(* IEC 61131-3 sources: JingjiangMoonbox/Application/Application/任务列表/TensionTask/电机运动/MotionCtl_GantryTrap/HandWheelCtl, 6 files *)

(* ---- StHandWheel.st ---- *)
(*@CES
Name=StHandWheel
Type=Gvl
TypeGuid=2db5746d-d284-4425-9f7f-2663a34b0ebc
Guid=e24024ef-b057-4603-89fd-c6f3dc30d212
HasDeclaration=True
HasImplementation=False
*)
{DECLARATION}
{attribute 'pack_mode' := '1'}
TYPE StHandWheel :
STRUCT
	wButton_HardWheel: WORD;(*手轮按键bit0-bit12对应按键1-13（手轮从左到右，从上到下）*)
// 	byRate_HardWheel: BYTE;(*倍率选择=13：X1;=14：X10;=15：X100;=16：X1000;=26：未定义（1000X后面还有一个档位）*)
// 	byAxisId_HardWheelCtl: BYTE;(*手轮旋钮当前选择
// 								=6：OFF
// 								=17：X
// 								=18：Y
// 								=19：Z
// 								=20：A*)

//2023.9.25.131020|手轮实际是倍率和轴选不是之前的定义，我们交换了一些2023.9.25.13110|
	byKnob_Right: BYTE;(*右选择=13：0档位;
								=14：1档位;
								=15：2档位;
								=16：3档位;
								=26：4档位（1000X后面还有一个档位）*)
	byKnob_Left: BYTE;(*左旋钮当前选择
								=6：0档位
								=17：1档位
								=18：2档位
								=19：3档位
								=20：4档位*)
	lrTargetPos_HardWheel: LREAL;(*当前手轮值-可以通过GT_RN_ZeroHandPos指令清除*)
	byHandWheelSts: BYTE;(**)
	asDisplay_HardWheel_HMI: ARRAY [1..4] OF STRING(16);(*手轮HMI显示-*)
	(*屏显功能说明：
	1.显示信号、电池电量
	2.当前操作色组号、当前操作的轴、标定模式以及标定轴、步进值
	3.显示版辊两侧电机实时位置(mm)
	4.显示网辊两侧电机实时位置(mm)
	(屏显格式说明：1行显示11个字符
	2/3/4行能显示16个字符)*)
	//2024.3.13.142250用于通讯给从站的变量
	arPos_HandWheel: ARRAY [1..4] OF REAL;//4个压力电机位置版辊M-G，网辊M-G
	byCtlId_HandWheel: BYTE;
	byCtlSts_HandWheel: BYTE;
						(*
							bit0:锁定模式
							bit1:运行模式
							bit2:标定DEBUG
							bit3:急停
							bit4:报警
							bit5:版/网切换
							bit6:清零处理
			2025.04.02.144750
							bit7:切换色组
						*)
END_STRUCT
END_TYPE

{IMPLEMENTATION}

(* ---- StHandWheel_BtnCtl.st ---- *)
(*@CES
Name=StHandWheel_BtnCtl
Type=Gvl
TypeGuid=2db5746d-d284-4425-9f7f-2663a34b0ebc
Guid=b84cb397-2bed-4490-8555-fa94b8c7b26f
HasDeclaration=True
HasImplementation=False
*)
{DECLARATION}
TYPE StHandWheel_BtnCtl :
STRUCT
	xReq_Inch_Net: BOOL;//匀墨
	xReqSwitch_Calib: BOOL;
	xReq_Confirm_Adjust_PressDn: BOOL;//位置矫正
	lrPos_HandWheelChange: LREAL;//手轮变化量

	xReqMove_M: BOOL;
	xReqMove_G: BOOL;
	xReqMoveUp: BOOL;
	xReqMoveDn: BOOL;

	xAdjust_V_Up : BOOL;
	xAdjust_V_Dn : BOOL;
	xAdjust_H_M : BOOL;
	xAdjust_H_G : BOOL;

//下面是需要区分版辊压力、网棍压力、张带辊压力的
	axReqLoad_Unload: ARRAY [1..gc_iMax_PressureRoller_Unit] OF BOOL;
	axReqPress_Up: ARRAY [1..gc_iMax_PressureRoller_Unit] OF BOOL;
	axReqPress_Dn: ARRAY [1..gc_iMax_PressureRoller_Unit] OF BOOL;

	axReqMoveFor: ARRAY [1..gc_iMax_PressureRoller_Unit] OF BOOL;
	axReqMoveRev: ARRAY [1..gc_iMax_PressureRoller_Unit] OF BOOL;

	axReq_Confirm_Load_Unload: ARRAY [1..gc_iMax_PressureRoller_Unit] OF BOOL;
	axReq_Confirm_press_up: ARRAY [1..gc_iMax_PressureRoller_Unit] OF BOOL;
	axReq_Confirm_press_dn: ARRAY [1..gc_iMax_PressureRoller_Unit] OF BOOL;

	axFlag_Ctl_Roller_All: ARRAY [1..gc_iMax_PressureRoller_Unit] OF BOOL;//控制的是同进同退-版辊
	axFlag_Ctl_Roller_M: ARRAY [1..gc_iMax_PressureRoller_Unit] OF BOOL;
	axFlag_Ctl_Roller_G: ARRAY [1..gc_iMax_PressureRoller_Unit] OF BOOL;

END_STRUCT
END_TYPE

{IMPLEMENTATION}

(* ---- KS_FB_HandwheelCtl.st ---- *)
(*@CES
Name=KS_FB_HandwheelCtl
Type=FunctionBlock
TypeGuid=6f9dac99-8de1-4efc-8465-68ac443b7d08
Guid=2f871db0-86b8-4868-b4d6-3d54ec95653d
HasDeclaration=True
HasImplementation=True
*)
{DECLARATION}
FUNCTION_BLOCK KS_FB_HandwheelCtl
VAR_INPUT
	i_xEn: BOOL;
	i_byUnitNumMax: BYTE;//色组数
	i_pastStHandWheel: POINTER TO ARRAY [1..MAX_UNIT_NUM] OF StHandWheel;
	i_pastStHandWheel_BtnCtl: POINTER TO ARRAY [1..MAX_UNIT_NUM] OF StHandWheel_BtnCtl;

	i_pabyUnitId_Ctl: POINTER TO ARRAY [1..MAX_UNIT_NUM] OF BYTE;//每个手持器控制的色组，可调整
	i_xFlag_Stop: BOOL;//停机状态
	i_xDebugMode: BOOL;//调试模式
	i_paxNeedZeroPos:  POINTER TO ARRAY [1..MAX_UNIT_NUM] OF BOOL;//手轮计数清零标志
	i_paxFlag_Mode_Calid: POINTER TO ARRAY [1..MAX_UNIT_NUM] OF BOOL;//手持器标定标值
	i_paxFlag_LockHandwheel: POINTER TO ARRAY [1..MAX_UNIT_NUM] OF BOOL;//手持器suoding
	//i_paxFlag_Ctl_Prn: POINTER TO ARRAY [1..MAX_UNIT_NUM] OF BOOL;
	i_paxEn_HandWheel: POINTER TO  ARRAY [1..MAX_UNIT_NUM] OF BOOL;
	i_paxAdjust_Auto_V: POINTER TO  ARRAY [1..MAX_UNIT_NUM] OF BOOL;
	i_paxAdjust_Auto_H: POINTER TO  ARRAY [1..MAX_UNIT_NUM] OF BOOL;

	i_paxAcc_UnitId : POINTER TO  ARRAY [1..MAX_UNIT_NUM] OF BOOL;
END_VAR
VAR_OUTPUT
END_VAR
VAR
	iN: INT;
	iM: INT;
	iRtn : INT;
	xFlag_Handwheel_Unit_One: BOOL;//手持器与色组一对一标值
	axFlag_LockHandwheel: ARRAY [1..MAX_UNIT_NUM] OF BOOL;//手持器锁定标值
	xInit: BOOL:= FALSE;//初始化一些东西
	astStHandWheel_Rec: ARRAY [1..MAX_UNIT_NUM] OF StHandWheel;
	aiCtlStep_Handwheel: ARRAY [1..MAX_UNIT_NUM] OF INT;//手持器锁定标值
	aiCtlUnit_Handwheel: ARRAY [1..MAX_UNIT_NUM] OF INT;//手持器锁定标值
	iTemp:INT:=1;
	aiStartUnitId:ARRAY [1..MAX_UNIT_NUM] OF INT;//非一对一手持器，每个手持器控制的起始
	aiStopUnitId:ARRAY [1..MAX_UNIT_NUM] OF INT;//非一对一手持器，每个手持器控制的结束色组号
	axFlag_Mode_Calid: ARRAY [1..MAX_UNIT_NUM] OF BOOL;//手持器标定标值
	iTimeCnt_Lock:INT:= 600;//超过600个周期没操作，认为可以锁定手轮了防止误操作
	iTimeCnt_Lock_Init:INT:= 3429;//超过600个周期没操作(2分钟)，手轮初始化一次防止进入休眠
	aiCnt_Lock_Num: ARRAY [1..MAX_UNIT_NUM] OF INT;
	aiCnt_Lock_Num_Init: ARRAY [1..MAX_UNIT_NUM] OF INT;
	axFlag_Lock: ARRAY [1..MAX_UNIT_NUM,1..5] OF BOOL;//手轮无动作标志
	iUnitIdCtl: INT;
	aiCnt_LockBtn: ARRAY [1..MAX_UNIT_NUM] OF INT;
	iTimeCnt_LockBtn:INT:= 20;//超过20个周期没操作，认为可以锁定手轮了防止误操作
	afbAcc_AxisId: ARRAY [1..MAX_UNIT_NUM] OF R_TRIG;
	afbDec_AxisId: ARRAY [1..MAX_UNIT_NUM] OF R_TRIG;
	abyAxisId_handwheel: ARRAY [1..MAX_UNIT_NUM] OF BYTE;
	axEn_HandWheel: ARRAY [1..MAX_UNIT_NUM] OF BOOL;
	iK: INT;
	afbTRIG_Switch_Calib: ARRAY [1..MAX_UNIT_NUM] OF R_TRIG;
	fbKS_FB_HandwheelCtl_Reset : KS_FB_HandwheelCtl_Reset;
	xFlag_En_ModeCalib : BOOL;
//2024.12.05.170136 | bai.zy
	xHandWheelCtlSignalUnit : BOOL;
	iHandWheelCount : INT;

	aiAccCtlUnitId_Handwheel: ARRAY [1..MAX_UNIT_NUM] OF INT;//切换色组时手持器锁定的色组号
END_VAR

{IMPLEMENTATION}
IF i_xEn THEN
	IF (i_byUnitNumMax>=1 AND i_byUnitNumMax<= MAX_UNIT_NUM) AND
		i_pastStHandWheel<>0 AND
		i_pabyUnitId_Ctl<>0 AND
		i_pastStHandWheel_BtnCtl <> 0 AND
		i_paxNeedZeroPos <> 0 AND
		i_paxFlag_Mode_Calid <> 0 AND
		i_paxEn_HandWheel <> 0 AND
		i_paxAdjust_Auto_V <> 0 AND
		i_paxAdjust_Auto_H <> 0 THEN

	//	i_pastStHandWheel^[2] := i_pastStHandWheel^[3];
		IF NOT xInit THEN
			xInit:= TRUE;
			FOR iN:=1 TO MAX_UNIT_NUM BY 1 DO
				axFlag_LockHandwheel[iN]:= TRUE;
				axFlag_Mode_Calid[iN]:= FALSE;
				FOR iM:=1 TO 5 BY 1 DO
					axFlag_Lock[iN,iM]:= FALSE;//用于判断手持器无动作的标志
				END_FOR
				aiCtlUnit_Handwheel[iN]:= MAX_UNIT_NUM;
				axEn_HandWheel[iN]:= FALSE;
			END_FOR

		ELSE//初始化完成就可以处理其他了
//2024.3.13.141555
// axEn_HandWheel[1]:= TRUE;
// axEn_HandWheel[2]:= FALSE;
			iHandWheelCount := 0;
			FOR iN := 1 TO i_byUnitNumMax BY 1 DO
				axEn_HandWheel[iN] := i_paxEn_HandWheel^[iN];
				IF axEn_HandWheel[iN] THEN
					iHandWheelCount := iHandWheelCount + 1;
				END_IF
			END_FOR

			IF iHandWheelCount = i_byUnitNumMax THEN
				xHandWheelCtlSignalUnit := TRUE;
			ELSE
				xHandWheelCtlSignalUnit := FALSE;
			END_IF

			FOR iN:=1 TO MAX_UNIT_NUM BY 1 DO
				IF axFlag_LockHandwheel[iN]  OR (NOT axEn_HandWheel[iN]) THEN
					aiCtlStep_Handwheel[iN]:= 1;//锁定状态
				ELSE
					IF xFlag_En_ModeCalib THEN//标定模式2023.7.26.094141更新轴选旋钮，先这么试一下
						IF i_xFlag_Stop AND i_xDebugMode THEN
							axFlag_Mode_Calid[aiCtlUnit_Handwheel[iN]]:= TRUE;
						ELSE
							axFlag_Mode_Calid[aiCtlUnit_Handwheel[iN]]:= FALSE;
							xFlag_En_ModeCalib := FALSE;
						END_IF
 					ELSE
 						axFlag_Mode_Calid[aiCtlUnit_Handwheel[iN]]:= FALSE;
 					END_IF

					IF axFlag_Mode_Calid[aiCtlUnit_Handwheel[iN]] THEN
						aiCtlStep_Handwheel[iN]:= 2;//标定模式
					ELSE
						aiCtlStep_Handwheel[iN]:= 3;//运行模式
					END_IF
				END_IF

			END_FOR
			//换一下吧2024.3.13.132259循环手轮数不好处理

			FOR iN:=1 TO i_byUnitNumMax BY 1 DO
//			FOR iN:=1 TO i_byHandWheel_Num BY 1 DO
				IF i_pastStHandWheel^[iN].wButton_HardWheel=0 THEN//无按钮按下
					axFlag_Lock[iN,1]:= TRUE;
				ELSE
					axFlag_Lock[iN,1]:= FALSE;
				END_IF
				IF i_pastStHandWheel^[iN].byKnob_Left-astStHandWheel_Rec[iN].byKnob_Left=0 THEN//轴选未操作
					axFlag_Lock[iN,2]:= TRUE;
				ELSE
					axFlag_Lock[iN,2]:= FALSE;
				END_IF
				IF i_pastStHandWheel^[iN].byKnob_Right-astStHandWheel_Rec[iN].byKnob_Right=0 THEN//右旋钮无动作
					axFlag_Lock[iN,3]:= TRUE;
				ELSE
					axFlag_Lock[iN,3]:= FALSE;
				END_IF
				IF i_pastStHandWheel^[iN].lrTargetPos_HardWheel-astStHandWheel_Rec[iN].lrTargetPos_HardWheel=0 THEN//手轮无动作
					axFlag_Lock[iN,4]:= TRUE;
				ELSE
					axFlag_Lock[iN,4]:= FALSE;
				END_IF
				IF axFlag_Lock[iN,1] AND axFlag_Lock[iN,2] AND axFlag_Lock[iN,3] AND axFlag_Lock[iN,4] THEN//手轮本周期无动作
					aiCnt_Lock_Num[iN]:= aiCnt_Lock_Num[iN]+1;
					aiCnt_Lock_Num_Init[iN] := aiCnt_Lock_Num_Init[iN] +1;
					IF aiCnt_Lock_Num[iN]>=iTimeCnt_Lock THEN//手持器持续600周期无动作-20s-进入锁定状态
						axFlag_LockHandwheel[iN]:= TRUE;
						aiCnt_Lock_Num[iN] := 0;
					END_IF
					IF aiCnt_Lock_Num_Init[iN]>= iTimeCnt_Lock_Init THEN
;//						iRtn := GT_RN_UsbInit();
						aiCnt_Lock_Num_Init[iN] := 0;
					END_IF
				ELSE
					aiCnt_Lock_Num[iN]:= 0;
					aiCnt_Lock_Num_Init[iN] := 0;
				END_IF

			END_FOR

			FOR iN:=1 TO i_byUnitNumMax BY 1 DO
//			FOR iN:=1 TO i_byHandWheel_Num BY 1 DO
				IF axEn_HandWheel[iN] THEN
					iUnitIdCtl:= aiCtlUnit_Handwheel[iN];
					afbAcc_AxisId[iN](CLK:= i_pastStHandWheel^[iN].wButton_HardWheel.0);
					afbDec_AxisId[iN](CLK:= i_pastStHandWheel^[iN].wButton_HardWheel.1);
					IF abyAxisId_handwheel[iN]<>i_pastStHandWheel^[iN].byKnob_Right THEN
						i_paxNeedZeroPos^[iN]:= TRUE;
						astStHandWheel_Rec[iN].lrTargetPos_HardWheel:= 0;//手轮值清零-好处理
						i_pastStHandWheel^[iN].lrTargetPos_HardWheel:= 0;
					END_IF
					abyAxisId_handwheel[iN]:= i_pastStHandWheel^[iN].byKnob_Right;
					CASE aiCtlStep_Handwheel[iN] OF
						1: //手轮锁定，不允许操作
						//锁定后，所有按钮输入不响应
							IF NOT i_paxAcc_UnitId^[iN] THEN
								IF i_pastStHandWheel^[iN].wButton_HardWheel.0 AND i_pastStHandWheel^[iN].wButton_HardWheel.11 THEN
									//两个按钮同时按下，就认为需要解锁
									axFlag_LockHandwheel[iN]:= FALSE;//解锁
									i_paxNeedZeroPos^[iN]:= TRUE;
									astStHandWheel_Rec[iN].lrTargetPos_HardWheel:= 0;//手轮值清零-好处理
									i_pastStHandWheel^[iN].lrTargetPos_HardWheel:= 0;

								END_IF
							ELSE
								IF afbAcc_AxisId[iN].Q THEN//继续增加
									iUnitIdCtl:= iUnitIdCtl+1;
									FOR iK:=1 TO i_byUnitNumMax BY 1 DO
										IF axEn_HandWheel[iK] THEN
											IF iUnitIdCtl= aiCtlUnit_Handwheel[iK] OR iUnitIdCtl > i_byUnitNumMax THEN//不能与其他手轮冲突
												IF iUnitIdCtl+1 > i_byUnitNumMax THEN//2024.12.05.133431 | bai.zy | 双手轮冲突、超过两个要重新做
													iUnitIdCtl:= 1;
												ELSE
													iUnitIdCtl:= iUnitIdCtl+1;
												END_IF
											END_IF
										END_IF
									END_FOR
									IF iUnitIdCtl>i_byUnitNumMax THEN
										iUnitIdCtl:= 1;
									END_IF
	// 								i_paxAcc_UnitId^[iN] := FALSE;
	// 								axFlag_LockHandwheel[iN]:= FALSE;//解锁
									i_paxNeedZeroPos^[iN]:= TRUE;
									astStHandWheel_Rec[iN].lrTargetPos_HardWheel:= 0;//手轮值清零-好处理
									i_pastStHandWheel^[iN].lrTargetPos_HardWheel:= 0;

									aiCtlUnit_Handwheel[iN]:=iUnitIdCtl;
								ELSIF i_pastStHandWheel^[iN].wButton_HardWheel.1 THEN//确认
									iUnitIdCtl:= iUnitIdCtl+1;
									FOR iK:=1 TO i_byUnitNumMax BY 1 DO
										IF axEn_HandWheel[iK] THEN
											IF iUnitIdCtl= aiCtlUnit_Handwheel[iK] OR iUnitIdCtl > i_byUnitNumMax THEN//不能与其他手轮冲突
												IF iUnitIdCtl+1 > i_byUnitNumMax THEN//2024.12.05.133431 | bai.zy | 双手轮冲突、超过两个要重新做
													iUnitIdCtl:= 1;
												ELSE
													iUnitIdCtl:= iUnitIdCtl+1;
												END_IF
											END_IF
										END_IF
									END_FOR
									IF iUnitIdCtl>i_byUnitNumMax THEN
										iUnitIdCtl:= 1;
									END_IF
									i_paxAcc_UnitId^[iN] := FALSE;
									axFlag_LockHandwheel[iN]:= FALSE;//解锁
									i_paxNeedZeroPos^[iN]:= TRUE;
									astStHandWheel_Rec[iN].lrTargetPos_HardWheel:= 0;//手轮值清零-好处理
									i_pastStHandWheel^[iN].lrTargetPos_HardWheel:= 0;

									IF xHandWheelCtlSignalUnit THEN
										aiCtlUnit_Handwheel[iN]:=iN;
									ELSE
										aiCtlUnit_Handwheel[iN]:=iUnitIdCtl;
									END_IF

								ELSIF i_pastStHandWheel^[iN].wButton_HardWheel.2 THEN//取消
									aiCtlUnit_Handwheel[iN] := aiAccCtlUnitId_Handwheel[iN];
									i_paxAcc_UnitId^[iN] := FALSE;
									axFlag_LockHandwheel[iN]:= FALSE;//解锁
									i_paxNeedZeroPos^[iN]:= TRUE;
									astStHandWheel_Rec[iN].lrTargetPos_HardWheel:= 0;//手轮值清零-好处理
									i_pastStHandWheel^[iN].lrTargetPos_HardWheel:= 0;
								ELSE//其他按键无效
									;
								END_IF
							END_IF

							afbTRIG_Switch_Calib[iN](CLK:= g_xModeCalibSwitch);
							g_xModeCalibSwitch := FALSE;
							IF afbTRIG_Switch_Calib[iN].Q THEN
								//axFlag_Mode_Calid[iUnitIdCtl]:= NOT axFlag_Mode_Calid[iUnitIdCtl];
								xFlag_En_ModeCalib:= NOT xFlag_En_ModeCalib;
							END_IF
		(*
		xReqMoveLeft: BOOL;
		xReqMoveRight: BOOL;
		xReqMoveUp: BOOL;
		xReqMoveDn: BOOL;
		xReqLoad_Unload: BOOL;
		xReqPress_Up: BOOL;
		xReqPress_Dn: BOOL;
		xReqSwitch_P_N: BOOL;
		xReqMoveFor: BOOL;
		xReqMoveRev: BOOL;
		xReq_Confirm_Load_Unload: BOOL;//
		xReq_Confirm_Load_Unload
		xReq_Confirm_press_up: BOOL;
		xReq_Confirm_press_dn: BOOL;
		*)
							i_pastStHandWheel_BtnCtl^[iUnitIdCtl].xReqMove_M:= FALSE;
							i_pastStHandWheel_BtnCtl^[iUnitIdCtl].xReqMove_G:= FALSE;
							i_pastStHandWheel_BtnCtl^[iUnitIdCtl].xReqMoveUp:= FALSE;
							i_pastStHandWheel_BtnCtl^[iUnitIdCtl].xReqMoveDn:= FALSE;
							i_pastStHandWheel_BtnCtl^[iUnitIdCtl].xReqSwitch_Calib:= FALSE;

							FOR iM :=1 TO gc_iMax_PressureRoller_Unit BY 1 DO
								i_pastStHandWheel_BtnCtl^[iUnitIdCtl].axReqLoad_Unload[iM]:= FALSE;
								i_pastStHandWheel_BtnCtl^[iUnitIdCtl].axReqPress_Up[iM]:= FALSE;
								i_pastStHandWheel_BtnCtl^[iUnitIdCtl].axReqPress_Dn[iM]:= FALSE;
								i_pastStHandWheel_BtnCtl^[iUnitIdCtl].axReqMoveFor[iM]:= FALSE;
								i_pastStHandWheel_BtnCtl^[iUnitIdCtl].axReqMoveRev[iM]:= FALSE;
								i_pastStHandWheel_BtnCtl^[iUnitIdCtl].axReq_Confirm_Load_Unload[iM]:= FALSE;
								i_pastStHandWheel_BtnCtl^[iUnitIdCtl].axReq_Confirm_press_up[iM]:= FALSE;
								i_pastStHandWheel_BtnCtl^[iUnitIdCtl].axReq_Confirm_press_dn[iM]:= FALSE;
							END_FOR

						2://标定模式
							IF afbAcc_AxisId[iN].Q THEN
								i_paxAcc_UnitId^[iN] := TRUE;
								aiAccCtlUnitId_Handwheel[iN] := iUnitIdCtl;
								axFlag_LockHandwheel[iN]:= TRUE;//锁定
								i_paxNeedZeroPos^[iN]:= TRUE;
								astStHandWheel_Rec[iN].lrTargetPos_HardWheel:= 0;//手轮值清零-好处理
								i_pastStHandWheel^[iN].lrTargetPos_HardWheel:= 0;
	// 							iUnitIdCtl:= iUnitIdCtl+1;
	// 							FOR iK:=1 TO i_byUnitNumMax BY 1 DO
	// 								IF axEn_HandWheel[iK] THEN
	// 									IF iUnitIdCtl= aiCtlUnit_Handwheel[iK] OR iUnitIdCtl > i_byUnitNumMax THEN//不能与其他手轮冲突
	// 										IF iUnitIdCtl+1 > i_byUnitNumMax THEN//2024.12.05.133431 | bai.zy | 双手轮冲突、超过两个要重新做
	// 											iUnitIdCtl:= 1;
	// 										ELSE
	// 											iUnitIdCtl:= iUnitIdCtl+1;
	// 										END_IF
	// 									END_IF
	// 								END_IF
	// 							END_FOR
	// 							IF iUnitIdCtl>i_byUnitNumMax THEN
	// 								iUnitIdCtl:= 1;
	// 							END_IF
	// 							i_paxNeedZeroPos^[iN]:= TRUE;
	// 							astStHandWheel_Rec[iN].lrTargetPos_HardWheel:= 0;//手轮值清零-好处理
	// 							i_pastStHandWheel^[iN].lrTargetPos_HardWheel:= 0;
	//
							END_IF//循环切换
	// 						IF xHandWheelCtlSignalUnit THEN
	// 							aiCtlUnit_Handwheel[iN]:=iN;
	// 						ELSE
	// 							aiCtlUnit_Handwheel[iN]:=iUnitIdCtl;
	// 						END_IF

							IF i_pastStHandWheel^[iN].byKnob_Left=18 THEN

								i_pastStHandWheel_BtnCtl^[iUnitIdCtl].axReq_Confirm_Load_Unload[1]:= i_pastStHandWheel^[iN].wButton_HardWheel.2;
								i_pastStHandWheel_BtnCtl^[iUnitIdCtl].axReq_Confirm_press_up[1]:= i_pastStHandWheel^[iN].wButton_HardWheel.5;
								i_pastStHandWheel_BtnCtl^[iUnitIdCtl].axReq_Confirm_press_dn[1]:= i_pastStHandWheel^[iN].wButton_HardWheel.9;

								i_pastStHandWheel_BtnCtl^[iUnitIdCtl].axFlag_Ctl_Roller_All[1]:=
									i_pastStHandWheel^[iN].byKnob_Right=13;
								i_pastStHandWheel_BtnCtl^[iUnitIdCtl].axFlag_Ctl_Roller_M[1]:=
									i_pastStHandWheel^[iN].byKnob_Right=14;
								i_pastStHandWheel_BtnCtl^[iUnitIdCtl].axFlag_Ctl_Roller_G[1]:=
									i_pastStHandWheel^[iN].byKnob_Right=15;
		//前进后退需要服用
								i_pastStHandWheel_BtnCtl^[iUnitIdCtl].axReqMoveFor[1]:= i_pastStHandWheel^[iN].wButton_HardWheel.7;
								i_pastStHandWheel_BtnCtl^[iUnitIdCtl].axReqMoveRev[1]:= i_pastStHandWheel^[iN].wButton_HardWheel.8;
								fbKS_FB_HandwheelCtl_Reset(i_iD:= 2, i_pstStHandWheel_BtnCtl:= ADR(i_pastStHandWheel_BtnCtl^[iUnitIdCtl]));
								fbKS_FB_HandwheelCtl_Reset(i_iD:= 3, i_pstStHandWheel_BtnCtl:= ADR(i_pastStHandWheel_BtnCtl^[iUnitIdCtl]));
							ELSIF i_pastStHandWheel^[iN].byKnob_Left=19 THEN
								i_pastStHandWheel_BtnCtl^[iUnitIdCtl].axReq_Confirm_Load_Unload[2]:= i_pastStHandWheel^[iN].wButton_HardWheel.2;
								i_pastStHandWheel_BtnCtl^[iUnitIdCtl].axReq_Confirm_press_up[2]:= i_pastStHandWheel^[iN].wButton_HardWheel.5;
								i_pastStHandWheel_BtnCtl^[iUnitIdCtl].axReq_Confirm_press_dn[2]:= i_pastStHandWheel^[iN].wButton_HardWheel.9;

								i_pastStHandWheel_BtnCtl^[iUnitIdCtl].axFlag_Ctl_Roller_All[2]:=
									i_pastStHandWheel^[iN].byKnob_Right=13;
								i_pastStHandWheel_BtnCtl^[iUnitIdCtl].axFlag_Ctl_Roller_M[2]:=
									i_pastStHandWheel^[iN].byKnob_Right=14;
								i_pastStHandWheel_BtnCtl^[iUnitIdCtl].axFlag_Ctl_Roller_G[2]:=
									i_pastStHandWheel^[iN].byKnob_Right=15;
		//前进后退需要服用
								i_pastStHandWheel_BtnCtl^[iUnitIdCtl].axReqMoveFor[2]:= i_pastStHandWheel^[iN].wButton_HardWheel.7;
								i_pastStHandWheel_BtnCtl^[iUnitIdCtl].axReqMoveRev[2]:= i_pastStHandWheel^[iN].wButton_HardWheel.8;
								fbKS_FB_HandwheelCtl_Reset(i_iD:= 1, i_pstStHandWheel_BtnCtl:= ADR(i_pastStHandWheel_BtnCtl^[iUnitIdCtl]));
								fbKS_FB_HandwheelCtl_Reset(i_iD:= 3, i_pstStHandWheel_BtnCtl:= ADR(i_pastStHandWheel_BtnCtl^[iUnitIdCtl]));
							ELSIF i_pastStHandWheel^[iN].byKnob_Left=20 THEN
								i_pastStHandWheel_BtnCtl^[iUnitIdCtl].axReq_Confirm_Load_Unload[3]:= i_pastStHandWheel^[iN].wButton_HardWheel.2;
								i_pastStHandWheel_BtnCtl^[iUnitIdCtl].axReq_Confirm_press_up[3]:= i_pastStHandWheel^[iN].wButton_HardWheel.5;
								i_pastStHandWheel_BtnCtl^[iUnitIdCtl].axReq_Confirm_press_dn[3]:= i_pastStHandWheel^[iN].wButton_HardWheel.9;

								i_pastStHandWheel_BtnCtl^[iUnitIdCtl].axFlag_Ctl_Roller_All[3]:=
									i_pastStHandWheel^[iN].byKnob_Right=13;
								i_pastStHandWheel_BtnCtl^[iUnitIdCtl].axFlag_Ctl_Roller_M[3]:=
									i_pastStHandWheel^[iN].byKnob_Right=14;
								i_pastStHandWheel_BtnCtl^[iUnitIdCtl].axFlag_Ctl_Roller_G[3]:=
									i_pastStHandWheel^[iN].byKnob_Right=15;
		//前进后退需要服用
								i_pastStHandWheel_BtnCtl^[iUnitIdCtl].axReqMoveFor[3]:= i_pastStHandWheel^[iN].wButton_HardWheel.7;
								i_pastStHandWheel_BtnCtl^[iUnitIdCtl].axReqMoveRev[3]:= i_pastStHandWheel^[iN].wButton_HardWheel.8;
								fbKS_FB_HandwheelCtl_Reset(i_iD:= 1, i_pstStHandWheel_BtnCtl:= ADR(i_pastStHandWheel_BtnCtl^[iUnitIdCtl]));
								fbKS_FB_HandwheelCtl_Reset(i_iD:= 2, i_pstStHandWheel_BtnCtl:= ADR(i_pastStHandWheel_BtnCtl^[iUnitIdCtl]));
							ELSE
								FOR iM := 1 TO gc_iMax_PressureRoller_Unit BY 1 DO
									fbKS_FB_HandwheelCtl_Reset(i_iD:= iM, i_pstStHandWheel_BtnCtl:= ADR(i_pastStHandWheel_BtnCtl^[iUnitIdCtl]));
								END_FOR
							END_IF

							afbTRIG_Switch_Calib[iN](CLK:= i_pastStHandWheel^[iN].wButton_HardWheel.12 OR g_xModeCalibSwitch);
							g_xModeCalibSwitch := FALSE;
							IF afbTRIG_Switch_Calib[iN].Q THEN
								//axFlag_Mode_Calid[iUnitIdCtl]:= NOT axFlag_Mode_Calid[iUnitIdCtl];
								xFlag_En_ModeCalib:= NOT xFlag_En_ModeCalib;
							END_IF

							IF i_pastStHandWheel^[iN].wButton_HardWheel= 2048 THEN//单独按下锁定才生效
								aiCnt_LockBtn[iN]:= aiCnt_LockBtn[iN]+1;
								IF aiCnt_LockBtn[iN]>iTimeCnt_LockBtn THEN
									axFlag_LockHandwheel[iN]:= TRUE;
								END_IF
							ELSE
								aiCnt_LockBtn[iN]:= 0;
							END_IF
							i_pastStHandWheel_BtnCtl^[iUnitIdCtl].lrPos_HandWheelChange:= i_pastStHandWheel^[iN].lrTargetPos_HardWheel-
										astStHandWheel_Rec[iN].lrTargetPos_HardWheel;
						3://运行模式
							IF afbAcc_AxisId[iN].Q THEN
								i_paxAcc_UnitId^[iN] := TRUE;
								aiAccCtlUnitId_Handwheel[iN] := iUnitIdCtl;
								axFlag_LockHandwheel[iN]:= TRUE;//锁定
								i_paxNeedZeroPos^[iN]:= TRUE;
								astStHandWheel_Rec[iN].lrTargetPos_HardWheel:= 0;//手轮值清零-好处理
								i_pastStHandWheel^[iN].lrTargetPos_HardWheel:= 0;
	// 							iUnitIdCtl:= iUnitIdCtl+1;
	// 							FOR iK:=1 TO i_byUnitNumMax BY 1 DO
	// 								IF axEn_HandWheel[iK] THEN
	// 									IF iUnitIdCtl= aiCtlUnit_Handwheel[iK] OR iUnitIdCtl > i_byUnitNumMax THEN//不能与其他手轮冲突
	// 										IF iUnitIdCtl+1 > i_byUnitNumMax THEN//2024.12.05.133431 | bai.zy | 双手轮冲突、超过两个要重新做
	// 											iUnitIdCtl:= 1;
	// 										ELSE
	// 											iUnitIdCtl:= iUnitIdCtl+1;
	// 										END_IF
	// 									END_IF
	// 								END_IF
	// 							END_FOR
	// 							IF iUnitIdCtl>i_byUnitNumMax THEN
	// 								iUnitIdCtl:= 1;
	// 							END_IF
	// 							i_paxNeedZeroPos^[iN]:= TRUE;
	// 							astStHandWheel_Rec[iN].lrTargetPos_HardWheel:= 0;//手轮值清零-好处理
	// 							i_pastStHandWheel^[iN].lrTargetPos_HardWheel:= 0;
	//
							END_IF
	// 						IF xHandWheelCtlSignalUnit THEN
	// 							aiCtlUnit_Handwheel[iN]:=iN;
	// 						ELSE
	// 							aiCtlUnit_Handwheel[iN]:=iUnitIdCtl;
	// 						END_IF

							IF i_pastStHandWheel^[iN].byKnob_Left=18 THEN
								i_pastStHandWheel_BtnCtl^[iUnitIdCtl].axReqLoad_Unload[1]:= i_pastStHandWheel^[iN].wButton_HardWheel.2 AND i_pastStHandWheel^[iN].wButton_HardWheel.11;
								i_pastStHandWheel_BtnCtl^[iUnitIdCtl].axReqPress_Up[1]:= i_pastStHandWheel^[iN].wButton_HardWheel.5 AND i_pastStHandWheel^[iN].wButton_HardWheel.11;
								i_pastStHandWheel_BtnCtl^[iUnitIdCtl].axReqPress_Dn[1]:= i_pastStHandWheel^[iN].wButton_HardWheel.9 AND i_pastStHandWheel^[iN].wButton_HardWheel.11;

								i_pastStHandWheel_BtnCtl^[iUnitIdCtl].axFlag_Ctl_Roller_All[1]:=
									i_pastStHandWheel^[iN].byKnob_Right=13;
								i_pastStHandWheel_BtnCtl^[iUnitIdCtl].axFlag_Ctl_Roller_M[1]:=
									i_pastStHandWheel^[iN].byKnob_Right=14;
								i_pastStHandWheel_BtnCtl^[iUnitIdCtl].axFlag_Ctl_Roller_G[1]:=
									i_pastStHandWheel^[iN].byKnob_Right=15;
								fbKS_FB_HandwheelCtl_Reset(i_iD:= 3, i_pstStHandWheel_BtnCtl:= ADR(i_pastStHandWheel_BtnCtl^[iUnitIdCtl]));
								fbKS_FB_HandwheelCtl_Reset(i_iD:= 2, i_pstStHandWheel_BtnCtl:= ADR(i_pastStHandWheel_BtnCtl^[iUnitIdCtl]));
							ELSIF i_pastStHandWheel^[iN].byKnob_Left=19 THEN
								i_pastStHandWheel_BtnCtl^[iUnitIdCtl].axReqLoad_Unload[2]:= i_pastStHandWheel^[iN].wButton_HardWheel.2 AND i_pastStHandWheel^[iN].wButton_HardWheel.11;
								i_pastStHandWheel_BtnCtl^[iUnitIdCtl].axReqPress_Up[2]:= i_pastStHandWheel^[iN].wButton_HardWheel.5 AND i_pastStHandWheel^[iN].wButton_HardWheel.11;
								i_pastStHandWheel_BtnCtl^[iUnitIdCtl].axReqPress_Dn[2]:= i_pastStHandWheel^[iN].wButton_HardWheel.9 AND i_pastStHandWheel^[iN].wButton_HardWheel.11;

								i_pastStHandWheel_BtnCtl^[iUnitIdCtl].axFlag_Ctl_Roller_All[2]:=
									i_pastStHandWheel^[iN].byKnob_Right=13;
								i_pastStHandWheel_BtnCtl^[iUnitIdCtl].axFlag_Ctl_Roller_M[2]:=
									i_pastStHandWheel^[iN].byKnob_Right=14;
								i_pastStHandWheel_BtnCtl^[iUnitIdCtl].axFlag_Ctl_Roller_G[2]:=
									i_pastStHandWheel^[iN].byKnob_Right=15;
								fbKS_FB_HandwheelCtl_Reset(i_iD:= 1, i_pstStHandWheel_BtnCtl:= ADR(i_pastStHandWheel_BtnCtl^[iUnitIdCtl]));
								fbKS_FB_HandwheelCtl_Reset(i_iD:= 3, i_pstStHandWheel_BtnCtl:= ADR(i_pastStHandWheel_BtnCtl^[iUnitIdCtl]));
							ELSIF i_pastStHandWheel^[iN].byKnob_Left=20 THEN
								i_pastStHandWheel_BtnCtl^[iUnitIdCtl].axReqLoad_Unload[3]:= i_pastStHandWheel^[iN].wButton_HardWheel.2 AND i_pastStHandWheel^[iN].wButton_HardWheel.11;
								i_pastStHandWheel_BtnCtl^[iUnitIdCtl].axReqPress_Up[3]:= i_pastStHandWheel^[iN].wButton_HardWheel.5 AND i_pastStHandWheel^[iN].wButton_HardWheel.11;
								i_pastStHandWheel_BtnCtl^[iUnitIdCtl].axReqPress_Dn[3]:= i_pastStHandWheel^[iN].wButton_HardWheel.9 AND i_pastStHandWheel^[iN].wButton_HardWheel.11;

								i_pastStHandWheel_BtnCtl^[iUnitIdCtl].axFlag_Ctl_Roller_All[3]:=
									i_pastStHandWheel^[iN].byKnob_Right=13;
								i_pastStHandWheel_BtnCtl^[iUnitIdCtl].axFlag_Ctl_Roller_M[3]:=
									i_pastStHandWheel^[iN].byKnob_Right=14;
								i_pastStHandWheel_BtnCtl^[iUnitIdCtl].axFlag_Ctl_Roller_G[3]:=
									i_pastStHandWheel^[iN].byKnob_Right=15;
								fbKS_FB_HandwheelCtl_Reset(i_iD:= 1, i_pstStHandWheel_BtnCtl:= ADR(i_pastStHandWheel_BtnCtl^[iUnitIdCtl]));
								fbKS_FB_HandwheelCtl_Reset(i_iD:= 2, i_pstStHandWheel_BtnCtl:= ADR(i_pastStHandWheel_BtnCtl^[iUnitIdCtl]));
							ELSE
								FOR iM := 1 TO gc_iMax_PressureRoller_Unit BY 1 DO
									fbKS_FB_HandwheelCtl_Reset(i_iD:= iM, i_pstStHandWheel_BtnCtl:= ADR(i_pastStHandWheel_BtnCtl^[iUnitIdCtl]));
								END_FOR
							END_IF

							//2025.03.04.154540 | 横向
							IF i_paxAdjust_Auto_H^[iUnitIdCtl] THEN
								i_pastStHandWheel_BtnCtl^[iUnitIdCtl].xAdjust_H_M:= i_pastStHandWheel^[iN].wButton_HardWheel.3;
								i_pastStHandWheel_BtnCtl^[iUnitIdCtl].xAdjust_H_G:= i_pastStHandWheel^[iN].wButton_HardWheel.4;
							ELSE
								i_pastStHandWheel_BtnCtl^[iUnitIdCtl].xReqMove_M:= i_pastStHandWheel^[iN].wButton_HardWheel.3;
								i_pastStHandWheel_BtnCtl^[iUnitIdCtl].xReqMove_G:= i_pastStHandWheel^[iN].wButton_HardWheel.4;
							END_IF
							//2025.03.04.154550| 纵向
							IF i_paxAdjust_Auto_V^[iUnitIdCtl] THEN//自动是修正量
								i_pastStHandWheel_BtnCtl^[iUnitIdCtl].xAdjust_V_Up:= i_pastStHandWheel^[iN].wButton_HardWheel.7;
								i_pastStHandWheel_BtnCtl^[iUnitIdCtl].xAdjust_V_Dn:= i_pastStHandWheel^[iN].wButton_HardWheel.8;
							ELSE//手动是调整量
								i_pastStHandWheel_BtnCtl^[iUnitIdCtl].xReqMoveUp:= i_pastStHandWheel^[iN].wButton_HardWheel.7;
								i_pastStHandWheel_BtnCtl^[iUnitIdCtl].xReqMoveDn:= i_pastStHandWheel^[iN].wButton_HardWheel.8;
							END_IF

							i_pastStHandWheel_BtnCtl^[iUnitIdCtl].xReq_Inch_Net:= i_pastStHandWheel^[iN].wButton_HardWheel.1;
							i_pastStHandWheel_BtnCtl^[iUnitIdCtl].xReq_Confirm_Adjust_PressDn:= i_pastStHandWheel^[iN].wButton_HardWheel.6;

							afbTRIG_Switch_Calib[iN](CLK:= i_pastStHandWheel^[iN].wButton_HardWheel.12 OR g_xModeCalibSwitch);
							g_xModeCalibSwitch := FALSE;
							IF afbTRIG_Switch_Calib[iN].Q THEN
								//axFlag_Mode_Calid[iUnitIdCtl]:= NOT axFlag_Mode_Calid[iUnitIdCtl];
								xFlag_En_ModeCalib:= NOT xFlag_En_ModeCalib;
							END_IF

	// 						IF i_xFlag_Stop THEN//运行模式时，停机状态下需要前进后退吗？，先按这个复用吧-两个键同时按下
	// 							i_pastStHandWheel_BtnCtl^[iUnitIdCtl].xReqMoveFor:=
	// 								i_pastStHandWheel^[iN].wButton_HardWheel.7 AND i_pastStHandWheel^[iN].wButton_HardWheel.11;
	// 							i_pastStHandWheel_BtnCtl^[iUnitIdCtl].xReqMoveRev:=
	// 								i_pastStHandWheel^[iN].wButton_HardWheel.8 AND i_pastStHandWheel^[iN].wButton_HardWheel.11;
	// 						ELSE//非停机状态就不给用前进后退了吧，就靠这个手轮或者进入退出使用了
	// 							i_pastStHandWheel_BtnCtl^[iUnitIdCtl].xReqMoveFor:= FALSE;
	// 							i_pastStHandWheel_BtnCtl^[iUnitIdCtl].xReqMoveRev:= FALSE;
	// 						END_IF
							IF i_pastStHandWheel^[iN].wButton_HardWheel= 2048 THEN//单独按下锁定才生效
								aiCnt_LockBtn[iN]:= aiCnt_LockBtn[iN]+1;
								IF aiCnt_LockBtn[iN]>iTimeCnt_LockBtn THEN
									axFlag_LockHandwheel[iN]:= TRUE;
								END_IF
							ELSE
								aiCnt_LockBtn[iN]:= 0;
							END_IF
							i_pastStHandWheel_BtnCtl^[iUnitIdCtl].lrPos_HandWheelChange:= i_pastStHandWheel^[iN].lrTargetPos_HardWheel-
										astStHandWheel_Rec[iN].lrTargetPos_HardWheel;
					END_CASE
					i_pabyUnitId_Ctl^[iN]:= INT_TO_BYTE(aiCtlUnit_Handwheel[iN]);
	//				i_paxFlag_Ctl_Prn^[iUnitIdCtl]:= axFlag_Ctl_Prn[iUnitIdCtl];
					i_paxFlag_Mode_Calid^[iUnitIdCtl]:= axFlag_Mode_Calid[iUnitIdCtl];//手持器标定标值
					i_paxFlag_LockHandwheel^[iN]:= axFlag_LockHandwheel[iN];//手持器suoding
				ELSE
					i_pastStHandWheel^[iN].byCtlSts_HandWheel.7:= FALSE;
				END_IF
			END_FOR

			sysmemcpy(ADR(astStHandWheel_Rec),i_pastStHandWheel,SIZEOF(astStHandWheel_Rec));
		END_IF
	END_IF
END_IF

(* ---- KS_FB_HandwheelCtl_Reset.st ---- *)
(*@CES
Name=KS_FB_HandwheelCtl_Reset
Type=FunctionBlock
TypeGuid=6f9dac99-8de1-4efc-8465-68ac443b7d08
Guid=166e6113-4ec8-46e9-b440-4c67f8b36266
HasDeclaration=True
HasImplementation=True
*)
{DECLARATION}
FUNCTION_BLOCK KS_FB_HandwheelCtl_Reset
VAR_INPUT
	i_iD : INT;
	i_pstStHandWheel_BtnCtl : POINTER TO StHandWheel_BtnCtl;
END_VAR
VAR_OUTPUT
END_VAR
VAR
END_VAR

{IMPLEMENTATION}
i_pstStHandWheel_BtnCtl^.axReq_Confirm_Load_Unload[i_iD]:= FALSE;
i_pstStHandWheel_BtnCtl^.axReq_Confirm_press_up[i_iD]:=FALSE;
i_pstStHandWheel_BtnCtl^.axReq_Confirm_press_dn[i_iD]:= FALSE;
i_pstStHandWheel_BtnCtl^.axFlag_Ctl_Roller_All[i_iD]:= FALSE;
i_pstStHandWheel_BtnCtl^.axFlag_Ctl_Roller_M[i_iD]:= FALSE;
i_pstStHandWheel_BtnCtl^.axFlag_Ctl_Roller_G[i_iD]:= FALSE;
i_pstStHandWheel_BtnCtl^.axReqMoveFor[i_iD]:= FALSE;
i_pstStHandWheel_BtnCtl^.axReqMoveRev[i_iD]:= FALSE;

(* ---- KS_FB_HandWheelRd.st ---- *)
(*@CES
Name=KS_FB_HandWheelRd
Type=FunctionBlock
TypeGuid=6f9dac99-8de1-4efc-8465-68ac443b7d08
Guid=56e9b8aa-8bae-4116-9277-461cb8a3efcc
HasDeclaration=True
HasImplementation=True
*)
{DECLARATION}
FUNCTION_BLOCK KS_FB_HandWheelRd
VAR_INPUT
	i_xEn: BOOL;
	i_pastStHandWheel: POINTER TO ARRAY [1..MAX_UNIT_NUM] OF StHandWheel;
END_VAR
VAR_OUTPUT
END_VAR
VAR
	iN: INT;
	iM : INT;
	iCountAddBlankNum : INT;
	iRtn : INT;
	iRtn_Read: INT;
	iRtn_Write: INT;
	stStHandPrm: StHandWheelPrm;
	iRtn_UnitId : INT;
	asDisplay_HardWheel_HMI: ARRAY [1..MAX_UNIT_NUM,1..4] OF STRING(16);(*手轮HMI显示-*)
	axRtnCmp_HMI : ARRAY[1..MAX_UNIT_NUM,1..4] OF BOOL;
	xInit : BOOL;
	sDisplay_HardWheel_HMI1: STRING(11);
	sDisplay_HardWheel_HMI2: STRING(16);
	sDisplay_HardWheel_HMI3: STRING(16);
	sDisplay_HardWheel_HMI4: STRING(16);
	sDisplay_HardWheel_HMIAll : STRING(59);
	iLenDisplay_HardWheel_HMI1 : INT;
	iLenDisplay_HardWheel_HMI2 : INT;
	iLenDisplay_HardWheel_HMI3 : INT;
	iLenDisplay_HardWheel_HMI4 : INT;
	iBlankNum1 : INT;
	iBlankNum2 : INT;
	iBlankNum3 : INT;
	iBlankNum4 : INT;

	tTimeError : TIME;
	tTimeError1 : TIME;
	mtargetPos : LREAL;
	tTempPos : TIME;
	tTempPos2 : TIME;

	enc1 : REAL;
	lrlastenc : REAL;
	tTemp : TIME;
	tTemp2 : TIME;
	tDelta1 : TIME;

	tTemp1:TIME;
	tDelta:TIME;
	xMoving,xStopping:BOOL;
	prfPos : LREAL;
	targetPos1 : DINT;
	lrlastpos:LREAL;
	a:BOOL:= FALSE;
	b: BOOL;
	delta11 : TIME;
	m_TarPos: REAL;
	prfvalue:LREAL;
	targetpos:LREAL;
	rtn : INT;
	rtn_Stop : INT;
	timeStart : TIME;
	timeEnd : TIME;
	arTarPos : ARRAY[1..10000] OF REAL;
	stimeDelta : ARRAY [1..10000] OF TIME;
	count : DINT;
	m_TarPos222 : LREAL;
	m_vel : LREAL;
	rtn_Update : INT;
	rtn_Vel : INT;
	abykeyNum_A : ARRAY[1..1000] OF BYTE;
	countKeyNum : INT;

	timeNow : TIME;
	udiRtn : UDINT;
	stTimestamp: SYSTIME;
	stSysTimedate: RTS_SYSTIMEDATE;(* RTS_SYSTIMEDATE *)
	nowtime:STRING;
	iKK : INT;
END_VAR

{IMPLEMENTATION}
IF NOT xInit THEN
	IF iRtn = 0 THEN
		xInit := TRUE;
	ELSE
		;
	END_IF
END_IF

FOR iN:=1 TO MAX_UNIT_NUM BY 1 DO
	IF iN = 1 THEN
		iRtn_Read:= GT_RN_GetHandPrm(ADR(stStHandPrm));
		IF iRtn_Read<>0 THEN(*读取失败-继续读取*)
			;
		ELSE(*处理读取的数据*)
			i_pastStHandWheel^[iN].wButton_HardWheel:= 0;
			IF stStHandPrm.keyNum_A<>0 THEN
				i_pastStHandWheel^[iN].wButton_HardWheel:=i_pastStHandWheel^[iN].wButton_HardWheel OR SHL(1,(stStHandPrm.keyNum_A-1));
			END_IF

			IF stStHandPrm.keyNum_B<>0 THEN
				i_pastStHandWheel^[iN].wButton_HardWheel:=i_pastStHandWheel^[iN].wButton_HardWheel OR SHL(1,(stStHandPrm.keyNum_B-1));
			END_IF
			i_pastStHandWheel^[iN].byKnob_Right:= stStHandPrm.rate;
			i_pastStHandWheel^[iN].byKnob_Left:= stStHandPrm.axisId;
			i_pastStHandWheel^[iN].lrTargetPos_HardWheel:=stStHandPrm.targetPos;
		END_IF
	END_IF
END_FOR

//
// //2023.8.21.152152
// IF count > 5000-1 THEN
// 	count := 1;
// END_IF
//
// IF g_astStHandWheel[1].lrTargetPos_HardWheel <> m_TarPos222 THEN
// 	timeStart := TIME();
// 	count := count + 1;
// 	arTarPos[count] := g_astStHandWheel[1].lrTargetPos_HardWheel - m_TarPos222;
// 	m_TarPos222 := g_astStHandWheel[1].lrTargetPos_HardWheel;
// 	stimeDelta [count] := timeStart-timeEnd;
// 	timeEnd := timeStart;
// END_IF
//
//
// IF countKeyNum > 1000-1 THEN
// 	countKeyNum := 1000-2;
// END_IF
// IF stStHandPrm.axisId = 6 THEN
// 	abykeyNum_A[countKeyNum] := stStHandPrm.keyNum_A;
// 	countKeyNum := countKeyNum +1;
// END_IF
//2023.8.21.152148*)
//m_vel := arTarPos[count] * 8388/200;
// 2023.07.20.234031
// IF g_xSetVelTemp THEN
// 	g_xSetVelTemp := FALSE;
// 	//rtn_Vel := GT_SetVel(profile:= 4, vel:= g_VelTemp, station_id:= 0);
// 	//rtn_Vel := GT_SetVel(profile:= 12, vel:= g_VelTemp, station_id:= 0);
// 	rtn_Vel := GT_SetVel(profile:= 20, vel:= g_VelTemp, station_id:= 0);
// 	//rtn_Update := GT_Update(mask:= SHL(WORD#1, 4-1),0);
// 	//rtn_Update := GT_Update(mask:= SHL(WORD#1, 12-1),0);
// 	//rtn_Update := GT_Update(mask:= SHL(DWORD#1, 20-1),0);
// END_IF
//2023.07.20.234033
(*
(*手轮显示，测试使用*)
		g_astStHandWheel[1].asDisplay_HardWheel_HMI[1] := '   KESAI';
		g_astStHandWheel[1].asDisplay_HardWheel_HMI[2] := BYTE_TO_STRING(g_astStHandWheel[1].byRate_HardWheel);
		g_astStHandWheel[1].asDisplay_HardWheel_HMI[3] := BYTE_TO_STRING(g_astStHandWheel[1].byAxisId_HardWheelCtl);
		g_astStHandWheel[1].asDisplay_HardWheel_HMI[4] := DINT_TO_STRING(g_astStHandWheel[1].diTargetPos_HardWheel);
*)
(*
//2023.8.21.151901
enc1 := g_astStWatch_Sts_display[10].rPos_Prf;
IF ABS(enc1-lrlastenc)<168 AND tTemp1 <> T#0MS THEN
	IF tTemp2=T#0MS THEN
		tTemp2:=TIME();
		tDelta1:=tTemp2-tTemp1;
		a := false;
	END_IF
ELSE
	tTemp2:=T#0MS;
END_IF
lrlastenc:=enc1;

prfPos := stStHandPrm.targetPos;//[1].lrTargetPos_HardWheel;//.targetPos;
IF ABS(prfPos-lrlastpos) < 3  AND  a = TRUE THEN
	IF tTemp1=T#0MS THEN
		tTemp1:=TIME();
		rtn := GT_GetPrfPos(
		profile:= 1,
		pValue:= ADR(prfvalue),
		count:= 1,
		pClock:= 0,
		station_id:= 51);
		targetpos := prfPos;
		//rtn_Vel := GT_SetVel(profile:= 5, vel:= 0, station_id:= 0);
		//rtn_Stop := GT_Stop(mask:= 24, option:= 24, station_id:= 0);
		IF b THEN
			b := FALSE;
			tTimeError1 := TIME();
			delta11 := tTimeError1-tTimeError;
		END_IF
	END_IF
ELSE
	tTemp1:=T#0MS;
END_IF

IF ABS(prfPos-lrlastpos) > 3 THEN
	a:= TRUE;
	IF NOT b THEN
		b := TRUE;
		tTimeError := TIME();
		m_TarPos := prfPos;
	END_IF

END_IF

lrlastpos:=prfPos;
*)

(* ---- KS_FB_HandWheelRd_Wr.st ---- *)
(*@CES
Name=KS_FB_HandWheelRd_Wr
Type=FunctionBlock
TypeGuid=6f9dac99-8de1-4efc-8465-68ac443b7d08
Guid=44523763-61a9-4779-9c1b-89e0f1500c64
HasDeclaration=True
HasImplementation=True
*)
{DECLARATION}
FUNCTION_BLOCK KS_FB_HandWheelRd_Wr
VAR_INPUT
	i_xEn: BOOL;
	i_pastStHandWheel: POINTER TO ARRAY [1..MAX_UNIT_NUM] OF StHandWheel;
END_VAR
VAR_OUTPUT
END_VAR
VAR
	iN: INT;
	iM : INT;
	iCountAddBlankNum : INT;
	iRtn : INT;
	iRtn_Read: INT;
	iRtn_Write: INT;
	stStHandPrm: StHandWheelPrm;
	iRtn_UnitId : INT;
	asDisplay_HardWheel_HMI: ARRAY [1..MAX_UNIT_NUM,1..4] OF STRING(16);(*手轮HMI显示-*)
	axRtnCmp_HMI : ARRAY[1..MAX_UNIT_NUM,1..4] OF BOOL;
	xInit : BOOL;
	sDisplay_HardWheel_HMI1: STRING(11);
	sDisplay_HardWheel_HMI2: STRING(16);
	sDisplay_HardWheel_HMI3: STRING(16);
	sDisplay_HardWheel_HMI4: STRING(16);
	sDisplay_HardWheel_HMIAll : STRING(59);
	iLenDisplay_HardWheel_HMI1 : INT;
	iLenDisplay_HardWheel_HMI2 : INT;
	iLenDisplay_HardWheel_HMI3 : INT;
	iLenDisplay_HardWheel_HMI4 : INT;
	iBlankNum1 : INT;
	iBlankNum2 : INT;
	iBlankNum3 : INT;
	iBlankNum4 : INT;

	tTimeError : TIME;
	tTimeError1 : TIME;
	mtargetPos : LREAL;
	tTempPos : TIME;
	tTempPos2 : TIME;

	enc1 : REAL;
	lrlastenc : REAL;
	tTemp : TIME;
	tTemp2 : TIME;
	tDelta1 : TIME;

	tTemp1:TIME;
	tDelta:TIME;
	xMoving,xStopping:BOOL;
	prfPos : LREAL;
	targetPos1 : DINT;
	lrlastpos:LREAL;
	a:BOOL:= FALSE;
	b: BOOL;
	delta11 : TIME;
	m_TarPos: REAL;
	prfvalue:LREAL;
	targetpos:LREAL;
	rtn : INT;
	rtn_Stop : INT;
	timeStart : TIME;
	timeEnd : TIME;
	arTarPos : ARRAY[1..10000] OF REAL;
	stimeDelta : ARRAY [1..10000] OF TIME;
	count : DINT;
	m_TarPos222 : LREAL;
	m_vel : LREAL;
	rtn_Update : INT;
	rtn_Vel : INT;
	abykeyNum_A : ARRAY[1..1000] OF BYTE;
	countKeyNum : INT;

	timeNow : TIME;
	udiRtn : UDINT;
	stTimestamp: SYSTIME;
	stSysTimedate: RTS_SYSTIMEDATE;(* RTS_SYSTIMEDATE *)
	nowtime:STRING;
	iKK : INT;
END_VAR

{IMPLEMENTATION}
IF NOT xInit THEN
	iRtn := GT_RN_UsbInit();
	IF iRtn = 0 THEN
		xInit := TRUE;
	ELSE
		;
	END_IF
END_IF

FOR iN:=1 TO MAX_UNIT_NUM BY 1 DO
	IF iN = 1 THEN
		sDisplay_HardWheel_HMI1 := i_pastStHandWheel^[iN].asDisplay_HardWheel_HMI[1];
		sDisplay_HardWheel_HMI2 := i_pastStHandWheel^[iN].asDisplay_HardWheel_HMI[2];
		sDisplay_HardWheel_HMI3 := i_pastStHandWheel^[iN].asDisplay_HardWheel_HMI[3];
		sDisplay_HardWheel_HMI4 := i_pastStHandWheel^[iN].asDisplay_HardWheel_HMI[4];
		iLenDisplay_HardWheel_HMI1 := LEN(sDisplay_HardWheel_HMI1);
		iLenDisplay_HardWheel_HMI2 := LEN(sDisplay_HardWheel_HMI2);
		iLenDisplay_HardWheel_HMI3 := LEN(sDisplay_HardWheel_HMI3);
		iLenDisplay_HardWheel_HMI4 := LEN(sDisplay_HardWheel_HMI4);
		iBlankNum1 := 11 - iLenDisplay_HardWheel_HMI1;
		iBlankNum2 := 16 - iLenDisplay_HardWheel_HMI2;
		iBlankNum3 := 16 - iLenDisplay_HardWheel_HMI3;
		iBlankNum4 := 16 - iLenDisplay_HardWheel_HMI4;
		FOR iCountAddBlankNum := 1 TO iBlankNum1 BY 1 DO
			sDisplay_HardWheel_HMI1 := CONCAT(sDisplay_HardWheel_HMI1,' ');
		END_FOR
		FOR iCountAddBlankNum := 1 TO iBlankNum2 BY 1 DO
			sDisplay_HardWheel_HMI2 := CONCAT(sDisplay_HardWheel_HMI2,' ');
		END_FOR
		FOR iCountAddBlankNum := 1 TO iBlankNum3 BY 1 DO
			sDisplay_HardWheel_HMI3 := CONCAT(sDisplay_HardWheel_HMI3,' ');
		END_FOR
		FOR iCountAddBlankNum := 1 TO iBlankNum4 BY 1 DO
			sDisplay_HardWheel_HMI4 := CONCAT(sDisplay_HardWheel_HMI4,' ');
		END_FOR
		sDisplay_HardWheel_HMIAll := sDisplay_HardWheel_HMI1;
		sDisplay_HardWheel_HMIAll := CONCAT(sDisplay_HardWheel_HMIAll,sDisplay_HardWheel_HMI2);
		sDisplay_HardWheel_HMIAll := CONCAT(sDisplay_HardWheel_HMIAll,sDisplay_HardWheel_HMI3);
		sDisplay_HardWheel_HMIAll := CONCAT(sDisplay_HardWheel_HMIAll,sDisplay_HardWheel_HMI4);
		iRtn:= GT_RN_Display(ADR(sDisplay_HardWheel_HMIAll));
	END_IF
END_FOR
